// TIA Portal V20 export
Screen "200APC1FX1Layout"  1276x673
  ScreenItem "Line_Header_X0_Y64" at 0,64 size 1276x0  Type=HmiLine
  ScreenItem "Title_ScreenOverview_X390_Y2" at 390,2 size 500x30  Type=HmiTextBox
  ScreenItem "permanentareaborderrectangle" at 0,0 size 0x0  Type=HmiRectangle
  ScreenItem "Button_Back" at 2,2 size 90x60  Type=HmiButton
  ScreenItem "Move_Legend" at 1184,2 size 90x60  Type=HmiButton
  ScreenItem "Fusszeile_Button_ManualOPMode1_2" at 188,2 size 90x60  Type=HmiButton
  ScreenItem "文本域_22" at 1107,604 size 104x23  Type=HmiTextBox
  ScreenItem "面板容器_23" at 1154,633 size 96x32  Type=HmiFaceplateContainer
  ScreenItem "面板容器_22" at 1049,633 size 96x32  Type=HmiFaceplateContainer
  ScreenItem "Fusszeile_Button_ManualOPMode1_1" at 95,2 size 90x60  Type=HmiButton
  ScreenItem "文本域_3" at 1133,87 size 93x23  Type=HmiTextBox
  ScreenItem "LSicar_Valve8Pos_LeftHomeRightWork_WithPB_5" at 1102,112 size 160x53  Type=HmiFaceplateContainer
  ScreenItem "文本域_1" at 1133,175 size 93x23  Type=HmiTextBox
  ScreenItem "LSicar_Valve8Pos_LeftHomeRightWork_WithPB_1" at 1102,200 size 160x53  Type=HmiFaceplateContainer
  ScreenItem "文本域_2" at 1132,263 size 93x23  Type=HmiTextBox
  ScreenItem "LSicar_Valve8Pos_LeftHomeRightWork_WithPB_2" at 1101,288 size 160x53  Type=HmiFaceplateContainer
  ScreenItem "文本域_5" at 1134,342 size 93x23  Type=HmiTextBox
  ScreenItem "LSicar_Valve8Pos_LeftHomeRightWork_WithPB_3" at 1103,367 size 160x53  Type=HmiFaceplateContainer
  ScreenItem "文本域_6" at 1134,430 size 93x23  Type=HmiTextBox
  ScreenItem "LSicar_Valve8Pos_LeftHomeRightWork_WithPB_4" at 1103,455 size 160x53  Type=HmiFaceplateContainer
  ScreenItem "文本域_7" at 1133,518 size 93x23  Type=HmiTextBox
  ScreenItem "LSicar_Valve8Pos_LeftHomeRightWork_WithPB_6" at 1102,543 size 160x53  Type=HmiFaceplateContainer
  ScreenItem "Graphic view_1" at 44,87 size 964x520  Type=HmiGraphicView
  ScreenItem "面板容器_24" at 1092,4 size 88x58  Type=HmiFaceplateContainer
  ScreenItem "OPMode1_Blocked" at 1166,6 size 14x14  Type=HmiGraphicView
  ScreenItem "OPMode4_Foreground_Blocked" at 1092,4 size 88x58  Type=HmiGraphicView
